(* IEC 61131-3 sources: llm-plc-st-eval/data/definitivo/claude-sonnet-4-6/I4/zero_shot, 3 files *)

(* ---- ejec_1.st ---- *)
```pascal
FUNCTION_BLOCK FB_EstrellaTriangulo
VAR_INPUT
    btnMarcha : BOOL; (* Pulsador de marcha *)
    btnParo   : BOOL; (* Pulsador de paro   *)
END_VAR

VAR_OUTPUT
    kM : BOOL; (* Contactor principal  *)
    kY : BOOL; (* Contactor estrella   *)
    kD : BOOL; (* Contactor triángulo  *)
END_VAR

VAR
    (* Temporizador para el tiempo en estrella: 8 s *)
    tEstrella  : TON;
    (* Temporizador para el tiempo muerto: 100 ms   *)
    tMuerto    : TON;

    (* Máquina de estados *)
    eEstado : INT;
    (*  0 = Reposo
        1 = Marcha en estrella
        2 = Tiempo muerto (kY abierto, kD aún cerrado)
        3 = Marcha en triángulo                        *)
END_VAR

(* ─────────────────────────────────────────────────────────────
   Lógica principal
   ───────────────────────────────────────────────────────────── *)

(* PARO: tiene prioridad absoluta en cualquier estado *)
IF btnParo THEN
    eEstado        := 0;
    tEstrella.IN   := FALSE;
    tMuerto.IN     := FALSE;
END_IF

CASE eEstado OF

    (* ── Estado 0: Reposo ─────────────────────────────────── *)
    0:
        kM := FALSE;
        kY := FALSE;
        kD := FALSE;

        IF btnMarcha AND NOT btnParo THEN
            eEstado := 1; (* Pasar a arranque en estrella *)
        END_IF

    (* ── Estado 1: Marcha en estrella ─────────────────────── *)
    1:
        kM := TRUE;
        kY := TRUE;  (* Estrella activa  *)
        kD := FALSE; (* Triángulo inactivo — nunca simultáneos *)

        (* Arrancar temporizador de 8 s *)
        tEstrella(IN := TRUE, PT := T#8S);

        IF tEstrella.Q THEN
            (* Tiempo en estrella cumplido: abrir kY *)
            tEstrella.IN := FALSE; (* Resetear temporizador *)
            eEstado      := 2;     (* Pasar a tiempo muerto  *)
        END_IF

    (* ── Estado 2: Tiempo muerto (100 ms) ─────────────────── *)
    2:
        kM := TRUE;
        kY := FALSE; (* Estrella ya desactivada  *)
        kD := FALSE; (* Triángulo aún inactivo   *)

        (* Arrancar temporizador de tiempo muerto *)
        tMuerto(IN := TRUE, PT := T#100MS);

        IF tMuerto.Q THEN
            (* Tiempo muerto cumplido: cerrar kD *)
            tMuerto.IN := FALSE; (* Resetear temporizador *)
            eEstado    := 3;     (* Pasar a marcha triángulo *)
        END_IF

    (* ── Estado 3: Marcha en triángulo ────────────────────── *)
    3:
        kM := TRUE;
        kY := FALSE; (* Estrella inactiva — nunca simultáneos *)
        kD := TRUE;  (* Triángulo activo *)

        (* Permanece aquí hasta que se pulse btnParo *)

    ELSE
        (* Estado desconocido: ir a reposo por seguridad *)
        eEstado := 0;

END_CASE

(* ─────────────────────────────────────────────────────────────
   Enclavamiento de seguridad hardware por software:
   garantizar que kY y kD nunca estén activos a la vez.
   ───────────────────────────────────────────────────────────── *)
IF kY AND kD THEN
    kY := FALSE;
    kD := FALSE;
    kM := FALSE;
    eEstado := 0; (* Volver a reposo ante condición anómala *)
END_IF
```

(* ---- ejec_2.st ---- *)
```pascal
FUNCTION_BLOCK FB_EstrellaTriangulo
VAR_INPUT
    btnMarcha : BOOL; (* Pulsador de marcha *)
    btnParo   : BOOL; (* Pulsador de paro   *)
END_VAR

VAR_OUTPUT
    kM : BOOL; (* Contactor principal  *)
    kY : BOOL; (* Contactor estrella   *)
    kD : BOOL; (* Contactor triángulo  *)
END_VAR

VAR
    (* Temporizador estrella: 8 s en estrella *)
    tEstrella  : TON;
    (* Temporizador tiempo muerto: 100 ms entre kY y kD *)
    tMuerto    : TON;

    (* Máquina de estados *)
    eEstado    : INT; (* 0=Reposo 1=Estrella 2=TiempoMuerto 3=Triangulo *)
END_VAR

(* ─────────────────────────────────────────────
   Lógica principal - Arranque Estrella-Triángulo
   ───────────────────────────────────────────── *)

(* PARO: tiene prioridad absoluta en cualquier estado *)
IF btnParo THEN
    eEstado := 0;
END_IF;

CASE eEstado OF

    (* ── Estado 0: Reposo ── *)
    0:
        kM := FALSE;
        kY := FALSE;
        kD := FALSE;
        tEstrella(IN := FALSE, PT := T#8S);    (* Resetear temporizadores *)
        tMuerto  (IN := FALSE, PT := T#100MS);

        IF btnMarcha AND NOT btnParo THEN
            eEstado := 1; (* Pasar a estrella *)
        END_IF;

    (* ── Estado 1: Funcionamiento en Estrella ── *)
    1:
        kM := TRUE;
        kY := TRUE;  (* Estrella activa  *)
        kD := FALSE; (* Triángulo inactivo - enclavamiento *)

        tEstrella(IN := TRUE, PT := T#8S);
        tMuerto  (IN := FALSE, PT := T#100MS); (* Mantener reseteado *)

        IF tEstrella.Q THEN
            kY      := FALSE;  (* Desactivar estrella antes de cambiar estado *)
            eEstado := 2;      (* Pasar a tiempo muerto *)
        END_IF;

    (* ── Estado 2: Tiempo Muerto (kY y kD ambos inactivos) ── *)
    2:
        kM := TRUE;
        kY := FALSE; (* Estrella inactiva  - enclavamiento garantizado *)
        kD := FALSE; (* Triángulo inactivo - enclavamiento garantizado *)

        tEstrella(IN := TRUE,  PT := T#8S);    (* Mantener Q activo para no resetear *)
        tMuerto  (IN := TRUE,  PT := T#100MS); (* Iniciar cuenta de tiempo muerto *)

        IF tMuerto.Q THEN
            eEstado := 3; (* Pasar a triángulo *)
        END_IF;

    (* ── Estado 3: Funcionamiento en Triángulo ── *)
    3:
        kM := TRUE;
        kY := FALSE; (* Estrella inactiva  - enclavamiento *)
        kD := TRUE;  (* Triángulo activo   *)

        tEstrella(IN := TRUE, PT := T#8S);    (* Mantener temporizadores estables *)
        tMuerto  (IN := TRUE, PT := T#100MS);

        (* Permanece en triángulo hasta que se pulse btnParo *)

    ELSE
        (* Estado desconocido: ir a reposo de forma segura *)
        eEstado := 0;

END_CASE;

(* Enclavamiento hardware por software: garantía adicional *)
(* kY y kD nunca pueden ser TRUE simultáneamente          *)
IF kY AND kD THEN
    kY := FALSE;
    kD := FALSE;
    kM := FALSE;
    eEstado := 0; (* Fallo: volver a reposo *)
END_IF;
```

(* ---- ejec_3.st ---- *)
```pascal
FUNCTION_BLOCK FB_EstrellaTriangulo
VAR_INPUT
    btnMarcha : BOOL; (* Pulsador de marcha *)
    btnParo   : BOOL; (* Pulsador de paro   *)
END_VAR

VAR_OUTPUT
    kM : BOOL; (* Contactor principal  *)
    kY : BOOL; (* Contactor estrella   *)
    kD : BOOL; (* Contactor triángulo  *)
END_VAR

VAR
    (* Temporizador para el tiempo en estrella: 8 s *)
    tEstrella  : TON;
    (* Temporizador para el tiempo muerto: 100 ms   *)
    tMuerto    : TON;

    (* Máquina de estados *)
    eEstado : INT := 0;
    (*
        0 = Reposo
        1 = Marcha en estrella
        2 = Tiempo muerto (kY y kD ambos OFF)
        3 = Marcha en triángulo
    *)
END_VAR

(* ─────────────────────────────────────────────────────────────
   Lógica principal: máquina de estados estrella-triángulo
   ───────────────────────────────────────────────────────────── *)

CASE eEstado OF

    (* ── Estado 0: Reposo ─────────────────────────────────── *)
    0:
        kM := FALSE;
        kY := FALSE;
        kD := FALSE;
        tEstrella(IN := FALSE, PT := T#8S);
        tMuerto  (IN := FALSE, PT := T#100MS);

        IF btnMarcha AND NOT btnParo THEN
            eEstado := 1; (* Pasar a arranque en estrella *)
        END_IF;

    (* ── Estado 1: Marcha en estrella ─────────────────────── *)
    1:
        kM := TRUE;
        kY := TRUE;  (* Estrella activa  *)
        kD := FALSE; (* Triángulo inactivo — interbloqueo *)

        (* Arrancar temporizador de estrella *)
        tEstrella(IN := TRUE, PT := T#8S);

        IF btnParo THEN
            eEstado := 0; (* Paro inmediato *)
        ELSIF tEstrella.Q THEN
            (* Tiempo en estrella cumplido → tiempo muerto *)
            tEstrella(IN := FALSE, PT := T#8S); (* Resetear *)
            eEstado := 2;
        END_IF;

    (* ── Estado 2: Tiempo muerto (100 ms) ─────────────────── *)
    2:
        kM := TRUE;
        kY := FALSE; (* Estrella ya desactivada  *)
        kD := FALSE; (* Triángulo aún inactivo   *)

        (* Arrancar temporizador de tiempo muerto *)
        tMuerto(IN := TRUE, PT := T#100MS);

        IF btnParo THEN
            eEstado := 0; (* Paro inmediato *)
        ELSIF tMuerto.Q THEN
            (* Tiempo muerto cumplido → activar triángulo *)
            tMuerto(IN := FALSE, PT := T#100MS); (* Resetear *)
            eEstado := 3;
        END_IF;

    (* ── Estado 3: Marcha en triángulo ────────────────────── *)
    3:
        kM := TRUE;
        kY := FALSE; (* Estrella inactiva — interbloqueo *)
        kD := TRUE;  (* Triángulo activo  *)

        IF btnParo THEN
            eEstado := 0; (* Paro inmediato *)
        END_IF;

    (* ── Estado por defecto: seguridad ───────────────────── *)
    ELSE
        eEstado := 0;

END_CASE;
```
